Fanuc KAREL source: KA00071.KL

PROGRAM KA00071
%NOLOCKGROUP
VAR
  SRC: XYZWPR
  DST: ARRAY[2] OF BYTE
BEGIN
  SRC.X = 1.0
  DST[1] = SRC
END KA00071
